(* IEC 61131-3 sources: codesys-to-astra/tests/POUs/FB_C2aStrings_Test, 8 files *)

(* ---- FB_C2aStrings_Test.decl.st ---- *)
// Назначение: набор тестов строковых замен OwenStringUtils (ожидания — по описанию ОВЕН v3.0, а не по коду).
// Автор:      kr0nsch
// Версия:     0.1.0
// Документ:   docs/TEST_REPORT.md
FUNCTION_BLOCK FB_C2aStrings_Test EXTENDS coUnit.FB_TestSuite
VAR CONSTANT
    R_DELTA : REAL := 0.0001;   // допуск сравнения REAL
END_VAR

(* ---- AddCharLeftRight.method.decl.st ---- *)
// ADD_CHAR дополняет слева и справа, длинную строку не меняет
METHOD PRIVATE AddCharLeftRight
VAR
    sL : STRING(255);  // слева
    sR : STRING(255);  // справа
    sLong : STRING(255);  // длиннее цели
END_VAR

(* ---- BeforeAfterFound.method.decl.st ---- *)
// Before/After по первому вхождению
METHOD PRIVATE BeforeAfterFound
VAR
    sB : STRING(255);  // Before
    sA : STRING(255);  // After
END_VAR

(* ---- BeforeAfterMissing.method.decl.st ---- *)
// подстрока не найдена — пустая строка
METHOD PRIVATE BeforeAfterMissing
VAR
    sB : STRING(255);  // Before
    sA : STRING(255);  // After
END_VAR

(* ---- Concat4.method.decl.st ---- *)
// CONCAT4 склеивает четыре строки
METHOD PRIVATE Concat4
VAR
    sResult : STRING(255);  // результат
END_VAR

(* ---- HexLowerNoPrefix.method.decl.st ---- *)
// WORD_TO_HEX_STR(16#BEEF, FALSE, '') = 'beef'
METHOD PRIVATE HexLowerNoPrefix
VAR
    sResult : STRING(8);  // результат
END_VAR

(* ---- HexStrRoundTrip.method.decl.st ---- *)
// HEX_STR_TO_WORD('0x1A2b', '0x') = 16#1A2B (регистр не важен)
METHOD PRIVATE HexStrRoundTrip
VAR
    wResult : WORD;  // результат
END_VAR

(* ---- HexUpperPadded.method.decl.st ---- *)
// WORD_TO_HEX_STR(16#00AF, TRUE, '0x') = '0x00AF' (допущение A9: 4 символа)
METHOD PRIVATE HexUpperPadded
VAR
    sResult : STRING(8);  // результат
END_VAR
